// TIA Portal V21 export
// export: Created 2026-10-09T20:27:06.6743102Z, ExportSetting WithDefaults, DisplayName Totally Integrated Automation Portal, DisplayVersion V21, DisplayName STEP 7 Professional, DisplayVersion V21, DisplayName STEP 7 Safety, DisplayVersion V21, DisplayName Tech WebApplication, DisplayVersion V21, DisplayName WinCC Basic/Comfort/Advanced, DisplayVersion V21, DisplayName WinCC Unified, DisplayVersion V21
FUNCTION_BLOCK "FB_Generate_Serial_Number"   // FB1, LAD
{ S7_Optimized_Access := 'TRUE' }
VERSION : 0.1
// stored: AutoNumber true, IsIECCheckEnabled false, IsRetainMemResEnabled false, MemoryReserve 100, SetENOAutomatically false, UDAEnableTagReadback false
   VAR_INPUT
      batchId : UDInt;
      productId : UDInt;
      productType : Int;
      trigger : Bool;
   END_VAR
   VAR_OUTPUT
      serialNumber : String;
      qrCode : USInt;
   END_VAR
   VAR
      sizeBatch : USInt;
      sizeId : USInt;
      retVal : USInt;
      dateString : String;
      batchString : String;
      productString : String;
      typeString : String;
      pTrigAux_1 : Bool;
   END_VAR
   VAR_TEMP
      localTime : DTL;
      qrNoTemp : String;
   END_VAR
   VAR_TEMP   // added for the SCL form of the ladder/FBD networks
      _w1 : Bool;
      _w2 : Bool;
   END_VAR
BEGIN

REGION Network 1 (SCL)
   // get string size of batch ID
   "FC_2_GetStringSizeOfNumber"(number:=#batchId,
                                stringSize=>#sizeBatch);

   // get string size of prodcut ID
   "FC_2_GetStringSizeOfNumber"(number:=#productId,
                                stringSize=>#sizeId);
END_REGION

REGION Network 2
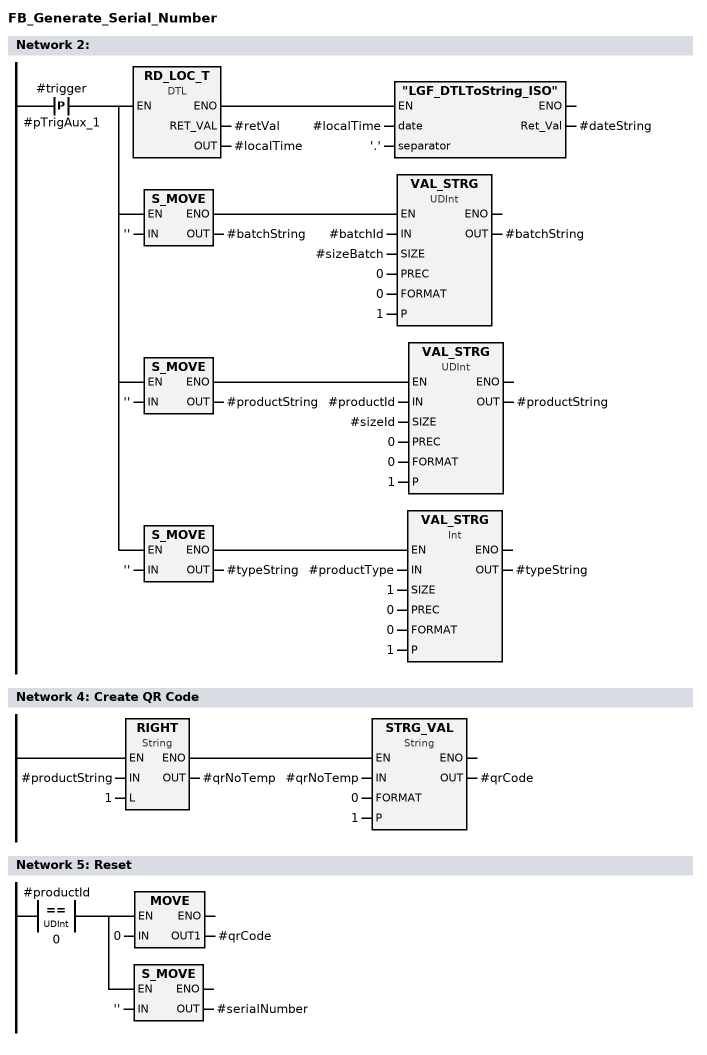
   RUNG wire#powerrail
      P_Contact(operand := #trigger, bit := #pTrigAux_1)
      wire#w1
      { S7_Templates := "date_type := DTL" } RD_LOC_T(RET_VAL => #retVal, OUT => #localTime)
      "LGF_DTLToString_ISO"("date" := #localTime, separator := '.', Ret_Val => #dateString)
   END_RUNG
   RUNG wire#w1
      S_Move(in := '', out => #batchString)
      { S7_Templates := "[value_type := UDInt, str_type := String]" } VAL_STRG(IN := #batchId, SIZE := #sizeBatch, PREC := 0, FORMAT := 0, P := 1, OUT => #batchString)
   END_RUNG
   RUNG wire#w1
      S_Move(in := '', out => #productString)
      { S7_Templates := "[value_type := UDInt, str_type := String]" } VAL_STRG(IN := #productId, SIZE := #sizeId, PREC := 0, FORMAT := 0, P := 1, OUT => #productString)
   END_RUNG
   RUNG wire#w1
      S_Move(in := '', out => #typeString)
      { S7_Templates := "[value_type := Int, str_type := String]" } VAL_STRG(IN := #productType, SIZE := 1, PREC := 0, FORMAT := 0, P := 1, OUT => #typeString)
   END_RUNG
   // the same network as SCL:
   #_w1 := #trigger AND NOT #pTrigAux_1;   // rising edge of #trigger
   #pTrigAux_1 := #trigger;
   #retVal := RD_LOC_T(EN := #_w1, OUT => #localTime, ENO => #_w2);
   IF #_w2 THEN #dateString := "LGF_DTLToString_ISO"("date" := #localTime, separator := '.'); END_IF;
   IF #_w1 THEN
       #batchString := '';
       VAL_STRG(IN := #batchId, SIZE := #sizeBatch, PREC := 0, FORMAT := 0, P := 1, OUT => #batchString);
       #productString := '';
       VAL_STRG(IN := #productId, SIZE := #sizeId, PREC := 0, FORMAT := 0, P := 1, OUT => #productString);
       #typeString := '';
       VAL_STRG(IN := #productType, SIZE := 1, PREC := 0, FORMAT := 0, P := 1, OUT => #typeString);
   END_IF;
END_REGION

REGION Network 3 (SCL): Create serial number
   #serialNumber := CONCAT(
                            IN1 := REPLACE(IN1:=DELETE(IN:=#dateString, L:=13, P:=17), IN2:='/', L:=1, P:=11),
                            IN2 := '/',
                            IN3 := #typeString,
                            IN4 := '/',
                            IN5 := #batchString,
                            IN6 := '/',
                            IN7 := #productString
   );
END_REGION

REGION Network 4: Create QR Code
   RUNG wire#powerrail
      { S7_Templates := "str_type := String" } RIGHT(IN := #productString, L := 1, OUT => #qrNoTemp)
      { S7_Templates := "[src_type := String, dest_type := USInt]" } STRG_VAL(IN := #qrNoTemp, FORMAT := 0, P := 1, OUT => #qrCode)
   END_RUNG
   // the same network as SCL:
   RIGHT(IN := #productString, L := 1, OUT => #qrNoTemp, ENO => #_w1);
   IF #_w1 THEN STRG_VAL(IN := #qrNoTemp, FORMAT := 0, P := 1, OUT => #qrCode); END_IF;
END_REGION

REGION Network 5: Reset
   RUNG wire#powerrail
      { S7_Templates := "SrcType := UDInt" } EQ_Contact(in1 := #productId, in2 := 0)
      wire#w1
      Move(in := 0, out1 => #qrCode)
   END_RUNG
   RUNG wire#w1
      S_Move(in := '', out => #serialNumber)
   END_RUNG
   // the same network as SCL:
   IF #productId = 0 THEN
       #qrCode := 0;
       #serialNumber := '';
   END_IF;
END_REGION
END_FUNCTION_BLOCK
